(* IEC 61131-3 sources: STAR-PLC-Agent/results/raw/batch_fresh_20261114/PUB007/functional/attempt_0001, 1 file *)

(* ---- test_program.st ---- *)
PROGRAM PLC_PRG
VAR
 BenchStep : UDINT := 0;
 BenchCalls : UDINT := 0;
 BenchDone : BOOL := FALSE;
 BenchUut0 : FB_Task;
 BenchUut1 : FB_Task;
 BenchUut2 : FB_Task;
 BenchUut3 : FB_Task;
 BenchUut4 : FB_Task;
 BenchUut5 : FB_Task;
 BenchUut6 : FB_Task;
 Binding_0_pumpGroup : ARRAY[1..5] OF ST_Pump;
 Binding_1_pumpGroup : ARRAY[1..5] OF ST_Pump;
 Binding_2_pumpGroup : ARRAY[1..5] OF ST_Pump;
 Binding_3_pumpGroup : ARRAY[1..5] OF ST_Pump;
 Binding_4_pumpGroup : ARRAY[1..5] OF ST_Pump;
 Binding_5_pumpGroup : ARRAY[1..5] OF ST_Pump;
 Binding_6_pumpGroup : ARRAY[1..5] OF ST_Pump;
 TraceIn_mode : ARRAY[0..29] OF BOOL;
 TraceIn_start : ARRAY[0..29] OF BOOL;
 TraceIn_stop : ARRAY[0..29] OF BOOL;
 TraceOut_pumpGroup_1_priority : ARRAY[0..29] OF INT;
 TraceOut_pumpGroup_1_selection : ARRAY[0..29] OF BOOL;
 TraceOut_pumpGroup_1_RunComd : ARRAY[0..29] OF BOOL;
 TraceOut_pumpGroup_2_priority : ARRAY[0..29] OF INT;
 TraceOut_pumpGroup_2_selection : ARRAY[0..29] OF BOOL;
 TraceOut_pumpGroup_2_RunComd : ARRAY[0..29] OF BOOL;
 TraceOut_pumpGroup_3_priority : ARRAY[0..29] OF INT;
 TraceOut_pumpGroup_3_selection : ARRAY[0..29] OF BOOL;
 TraceOut_pumpGroup_3_RunComd : ARRAY[0..29] OF BOOL;
 TraceOut_pumpGroup_4_priority : ARRAY[0..29] OF INT;
 TraceOut_pumpGroup_4_selection : ARRAY[0..29] OF BOOL;
 TraceOut_pumpGroup_4_RunComd : ARRAY[0..29] OF BOOL;
 TraceOut_pumpGroup_5_priority : ARRAY[0..29] OF INT;
 TraceOut_pumpGroup_5_selection : ARRAY[0..29] OF BOOL;
 TraceOut_pumpGroup_5_RunComd : ARRAY[0..29] OF BOOL;
END_VAR

IF NOT BenchDone THEN
 CASE BenchStep OF
 0:
   Binding_0_pumpGroup[1].priority := INT#10;
   Binding_0_pumpGroup[1].selection := TRUE;
   Binding_0_pumpGroup[1].RunComd := FALSE;
   Binding_0_pumpGroup[2].priority := INT#20;
   Binding_0_pumpGroup[2].selection := FALSE;
   Binding_0_pumpGroup[2].RunComd := FALSE;
   Binding_0_pumpGroup[3].priority := INT#30;
   Binding_0_pumpGroup[3].selection := TRUE;
   Binding_0_pumpGroup[3].RunComd := FALSE;
   Binding_0_pumpGroup[4].priority := INT#40;
   Binding_0_pumpGroup[4].selection := FALSE;
   Binding_0_pumpGroup[4].RunComd := FALSE;
   Binding_0_pumpGroup[5].priority := INT#50;
   Binding_0_pumpGroup[5].selection := FALSE;
   Binding_0_pumpGroup[5].RunComd := FALSE;
   BenchUut0.mode := FALSE;
   BenchUut0.start := TRUE;
   BenchUut0.stop := FALSE;
   TraceIn_mode[0] := BenchUut0.mode;
   TraceIn_start[0] := BenchUut0.start;
   TraceIn_stop[0] := BenchUut0.stop;
   BenchUut0(pumpGroup := Binding_0_pumpGroup);
   TraceOut_pumpGroup_1_priority[0] := Binding_0_pumpGroup[1].priority;
   TraceOut_pumpGroup_1_selection[0] := Binding_0_pumpGroup[1].selection;
   TraceOut_pumpGroup_1_RunComd[0] := Binding_0_pumpGroup[1].RunComd;
   TraceOut_pumpGroup_2_priority[0] := Binding_0_pumpGroup[2].priority;
   TraceOut_pumpGroup_2_selection[0] := Binding_0_pumpGroup[2].selection;
   TraceOut_pumpGroup_2_RunComd[0] := Binding_0_pumpGroup[2].RunComd;
   TraceOut_pumpGroup_3_priority[0] := Binding_0_pumpGroup[3].priority;
   TraceOut_pumpGroup_3_selection[0] := Binding_0_pumpGroup[3].selection;
   TraceOut_pumpGroup_3_RunComd[0] := Binding_0_pumpGroup[3].RunComd;
   TraceOut_pumpGroup_4_priority[0] := Binding_0_pumpGroup[4].priority;
   TraceOut_pumpGroup_4_selection[0] := Binding_0_pumpGroup[4].selection;
   TraceOut_pumpGroup_4_RunComd[0] := Binding_0_pumpGroup[4].RunComd;
   TraceOut_pumpGroup_5_priority[0] := Binding_0_pumpGroup[5].priority;
   TraceOut_pumpGroup_5_selection[0] := Binding_0_pumpGroup[5].selection;
   TraceOut_pumpGroup_5_RunComd[0] := Binding_0_pumpGroup[5].RunComd;
   BenchCalls := BenchCalls + 1;
 1:
   Binding_0_pumpGroup[1].priority := INT#10;
   Binding_0_pumpGroup[1].selection := TRUE;
   Binding_0_pumpGroup[1].RunComd := TRUE;
   Binding_0_pumpGroup[2].priority := INT#20;
   Binding_0_pumpGroup[2].selection := FALSE;
   Binding_0_pumpGroup[2].RunComd := FALSE;
   Binding_0_pumpGroup[3].priority := INT#30;
   Binding_0_pumpGroup[3].selection := TRUE;
   Binding_0_pumpGroup[3].RunComd := TRUE;
   Binding_0_pumpGroup[4].priority := INT#40;
   Binding_0_pumpGroup[4].selection := FALSE;
   Binding_0_pumpGroup[4].RunComd := FALSE;
   Binding_0_pumpGroup[5].priority := INT#50;
   Binding_0_pumpGroup[5].selection := FALSE;
   Binding_0_pumpGroup[5].RunComd := FALSE;
   BenchUut0.mode := FALSE;
   BenchUut0.start := FALSE;
   BenchUut0.stop := FALSE;
   TraceIn_mode[1] := BenchUut0.mode;
   TraceIn_start[1] := BenchUut0.start;
   TraceIn_stop[1] := BenchUut0.stop;
   BenchUut0(pumpGroup := Binding_0_pumpGroup);
   TraceOut_pumpGroup_1_priority[1] := Binding_0_pumpGroup[1].priority;
   TraceOut_pumpGroup_1_selection[1] := Binding_0_pumpGroup[1].selection;
   TraceOut_pumpGroup_1_RunComd[1] := Binding_0_pumpGroup[1].RunComd;
   TraceOut_pumpGroup_2_priority[1] := Binding_0_pumpGroup[2].priority;
   TraceOut_pumpGroup_2_selection[1] := Binding_0_pumpGroup[2].selection;
   TraceOut_pumpGroup_2_RunComd[1] := Binding_0_pumpGroup[2].RunComd;
   TraceOut_pumpGroup_3_priority[1] := Binding_0_pumpGroup[3].priority;
   TraceOut_pumpGroup_3_selection[1] := Binding_0_pumpGroup[3].selection;
   TraceOut_pumpGroup_3_RunComd[1] := Binding_0_pumpGroup[3].RunComd;
   TraceOut_pumpGroup_4_priority[1] := Binding_0_pumpGroup[4].priority;
   TraceOut_pumpGroup_4_selection[1] := Binding_0_pumpGroup[4].selection;
   TraceOut_pumpGroup_4_RunComd[1] := Binding_0_pumpGroup[4].RunComd;
   TraceOut_pumpGroup_5_priority[1] := Binding_0_pumpGroup[5].priority;
   TraceOut_pumpGroup_5_selection[1] := Binding_0_pumpGroup[5].selection;
   TraceOut_pumpGroup_5_RunComd[1] := Binding_0_pumpGroup[5].RunComd;
   BenchCalls := BenchCalls + 1;
 2:
   Binding_0_pumpGroup[1].priority := INT#10;
   Binding_0_pumpGroup[1].selection := TRUE;
   Binding_0_pumpGroup[1].RunComd := TRUE;
   Binding_0_pumpGroup[2].priority := INT#20;
   Binding_0_pumpGroup[2].selection := FALSE;
   Binding_0_pumpGroup[2].RunComd := FALSE;
   Binding_0_pumpGroup[3].priority := INT#30;
   Binding_0_pumpGroup[3].selection := TRUE;
   Binding_0_pumpGroup[3].RunComd := TRUE;
   Binding_0_pumpGroup[4].priority := INT#40;
   Binding_0_pumpGroup[4].selection := FALSE;
   Binding_0_pumpGroup[4].RunComd := FALSE;
   Binding_0_pumpGroup[5].priority := INT#50;
   Binding_0_pumpGroup[5].selection := FALSE;
   Binding_0_pumpGroup[5].RunComd := FALSE;
   BenchUut0.mode := FALSE;
   BenchUut0.start := TRUE;
   BenchUut0.stop := TRUE;
   TraceIn_mode[2] := BenchUut0.mode;
   TraceIn_start[2] := BenchUut0.start;
   TraceIn_stop[2] := BenchUut0.stop;
   BenchUut0(pumpGroup := Binding_0_pumpGroup);
   TraceOut_pumpGroup_1_priority[2] := Binding_0_pumpGroup[1].priority;
   TraceOut_pumpGroup_1_selection[2] := Binding_0_pumpGroup[1].selection;
   TraceOut_pumpGroup_1_RunComd[2] := Binding_0_pumpGroup[1].RunComd;
   TraceOut_pumpGroup_2_priority[2] := Binding_0_pumpGroup[2].priority;
   TraceOut_pumpGroup_2_selection[2] := Binding_0_pumpGroup[2].selection;
   TraceOut_pumpGroup_2_RunComd[2] := Binding_0_pumpGroup[2].RunComd;
   TraceOut_pumpGroup_3_priority[2] := Binding_0_pumpGroup[3].priority;
   TraceOut_pumpGroup_3_selection[2] := Binding_0_pumpGroup[3].selection;
   TraceOut_pumpGroup_3_RunComd[2] := Binding_0_pumpGroup[3].RunComd;
   TraceOut_pumpGroup_4_priority[2] := Binding_0_pumpGroup[4].priority;
   TraceOut_pumpGroup_4_selection[2] := Binding_0_pumpGroup[4].selection;
   TraceOut_pumpGroup_4_RunComd[2] := Binding_0_pumpGroup[4].RunComd;
   TraceOut_pumpGroup_5_priority[2] := Binding_0_pumpGroup[5].priority;
   TraceOut_pumpGroup_5_selection[2] := Binding_0_pumpGroup[5].selection;
   TraceOut_pumpGroup_5_RunComd[2] := Binding_0_pumpGroup[5].RunComd;
   BenchCalls := BenchCalls + 1;
 3:
   Binding_1_pumpGroup[1].priority := INT#10;
   Binding_1_pumpGroup[1].selection := TRUE;
   Binding_1_pumpGroup[1].RunComd := FALSE;
   Binding_1_pumpGroup[2].priority := INT#20;
   Binding_1_pumpGroup[2].selection := FALSE;
   Binding_1_pumpGroup[2].RunComd := FALSE;
   Binding_1_pumpGroup[3].priority := INT#30;
   Binding_1_pumpGroup[3].selection := TRUE;
   Binding_1_pumpGroup[3].RunComd := FALSE;
   Binding_1_pumpGroup[4].priority := INT#40;
   Binding_1_pumpGroup[4].selection := FALSE;
   Binding_1_pumpGroup[4].RunComd := FALSE;
   Binding_1_pumpGroup[5].priority := INT#50;
   Binding_1_pumpGroup[5].selection := FALSE;
   Binding_1_pumpGroup[5].RunComd := FALSE;
   BenchUut1.mode := TRUE;
   BenchUut1.start := TRUE;
   BenchUut1.stop := FALSE;
   TraceIn_mode[3] := BenchUut1.mode;
   TraceIn_start[3] := BenchUut1.start;
   TraceIn_stop[3] := BenchUut1.stop;
   BenchUut1(pumpGroup := Binding_1_pumpGroup);
   TraceOut_pumpGroup_1_priority[3] := Binding_1_pumpGroup[1].priority;
   TraceOut_pumpGroup_1_selection[3] := Binding_1_pumpGroup[1].selection;
   TraceOut_pumpGroup_1_RunComd[3] := Binding_1_pumpGroup[1].RunComd;
   TraceOut_pumpGroup_2_priority[3] := Binding_1_pumpGroup[2].priority;
   TraceOut_pumpGroup_2_selection[3] := Binding_1_pumpGroup[2].selection;
   TraceOut_pumpGroup_2_RunComd[3] := Binding_1_pumpGroup[2].RunComd;
   TraceOut_pumpGroup_3_priority[3] := Binding_1_pumpGroup[3].priority;
   TraceOut_pumpGroup_3_selection[3] := Binding_1_pumpGroup[3].selection;
   TraceOut_pumpGroup_3_RunComd[3] := Binding_1_pumpGroup[3].RunComd;
   TraceOut_pumpGroup_4_priority[3] := Binding_1_pumpGroup[4].priority;
   TraceOut_pumpGroup_4_selection[3] := Binding_1_pumpGroup[4].selection;
   TraceOut_pumpGroup_4_RunComd[3] := Binding_1_pumpGroup[4].RunComd;
   TraceOut_pumpGroup_5_priority[3] := Binding_1_pumpGroup[5].priority;
   TraceOut_pumpGroup_5_selection[3] := Binding_1_pumpGroup[5].selection;
   TraceOut_pumpGroup_5_RunComd[3] := Binding_1_pumpGroup[5].RunComd;
   BenchCalls := BenchCalls + 1;
 4:
   Binding_1_pumpGroup[1].priority := INT#5;
   Binding_1_pumpGroup[1].selection := TRUE;
   Binding_1_pumpGroup[1].RunComd := FALSE;
   Binding_1_pumpGroup[2].priority := INT#5;
   Binding_1_pumpGroup[2].selection := FALSE;
   Binding_1_pumpGroup[2].RunComd := FALSE;
   Binding_1_pumpGroup[3].priority := INT#5;
   Binding_1_pumpGroup[3].selection := TRUE;
   Binding_1_pumpGroup[3].RunComd := TRUE;
   Binding_1_pumpGroup[4].priority := INT#5;
   Binding_1_pumpGroup[4].selection := FALSE;
   Binding_1_pumpGroup[4].RunComd := TRUE;
   Binding_1_pumpGroup[5].priority := INT#5;
   Binding_1_pumpGroup[5].selection := FALSE;
   Binding_1_pumpGroup[5].RunComd := TRUE;
   BenchUut1.mode := TRUE;
   BenchUut1.start := TRUE;
   BenchUut1.stop := FALSE;
   TraceIn_mode[4] := BenchUut1.mode;
   TraceIn_start[4] := BenchUut1.start;
   TraceIn_stop[4] := BenchUut1.stop;
   BenchUut1(pumpGroup := Binding_1_pumpGroup);
   TraceOut_pumpGroup_1_priority[4] := Binding_1_pumpGroup[1].priority;
   TraceOut_pumpGroup_1_selection[4] := Binding_1_pumpGroup[1].selection;
   TraceOut_pumpGroup_1_RunComd[4] := Binding_1_pumpGroup[1].RunComd;
   TraceOut_pumpGroup_2_priority[4] := Binding_1_pumpGroup[2].priority;
   TraceOut_pumpGroup_2_selection[4] := Binding_1_pumpGroup[2].selection;
   TraceOut_pumpGroup_2_RunComd[4] := Binding_1_pumpGroup[2].RunComd;
   TraceOut_pumpGroup_3_priority[4] := Binding_1_pumpGroup[3].priority;
   TraceOut_pumpGroup_3_selection[4] := Binding_1_pumpGroup[3].selection;
   TraceOut_pumpGroup_3_RunComd[4] := Binding_1_pumpGroup[3].RunComd;
   TraceOut_pumpGroup_4_priority[4] := Binding_1_pumpGroup[4].priority;
   TraceOut_pumpGroup_4_selection[4] := Binding_1_pumpGroup[4].selection;
   TraceOut_pumpGroup_4_RunComd[4] := Binding_1_pumpGroup[4].RunComd;
   TraceOut_pumpGroup_5_priority[4] := Binding_1_pumpGroup[5].priority;
   TraceOut_pumpGroup_5_selection[4] := Binding_1_pumpGroup[5].selection;
   TraceOut_pumpGroup_5_RunComd[4] := Binding_1_pumpGroup[5].RunComd;
   BenchCalls := BenchCalls + 1;
 5:
   Binding_1_pumpGroup[1].priority := INT#-3;
   Binding_1_pumpGroup[1].selection := TRUE;
   Binding_1_pumpGroup[1].RunComd := TRUE;
   Binding_1_pumpGroup[2].priority := INT#0;
   Binding_1_pumpGroup[2].selection := FALSE;
   Binding_1_pumpGroup[2].RunComd := TRUE;
   Binding_1_pumpGroup[3].priority := INT#-1;
   Binding_1_pumpGroup[3].selection := TRUE;
   Binding_1_pumpGroup[3].RunComd := TRUE;
   Binding_1_pumpGroup[4].priority := INT#-2;
   Binding_1_pumpGroup[4].selection := FALSE;
   Binding_1_pumpGroup[4].RunComd := FALSE;
   Binding_1_pumpGroup[5].priority := INT#4;
   Binding_1_pumpGroup[5].selection := FALSE;
   Binding_1_pumpGroup[5].RunComd := FALSE;
   BenchUut1.mode := TRUE;
   BenchUut1.start := TRUE;
   BenchUut1.stop := FALSE;
   TraceIn_mode[5] := BenchUut1.mode;
   TraceIn_start[5] := BenchUut1.start;
   TraceIn_stop[5] := BenchUut1.stop;
   BenchUut1(pumpGroup := Binding_1_pumpGroup);
   TraceOut_pumpGroup_1_priority[5] := Binding_1_pumpGroup[1].priority;
   TraceOut_pumpGroup_1_selection[5] := Binding_1_pumpGroup[1].selection;
   TraceOut_pumpGroup_1_RunComd[5] := Binding_1_pumpGroup[1].RunComd;
   TraceOut_pumpGroup_2_priority[5] := Binding_1_pumpGroup[2].priority;
   TraceOut_pumpGroup_2_selection[5] := Binding_1_pumpGroup[2].selection;
   TraceOut_pumpGroup_2_RunComd[5] := Binding_1_pumpGroup[2].RunComd;
   TraceOut_pumpGroup_3_priority[5] := Binding_1_pumpGroup[3].priority;
   TraceOut_pumpGroup_3_selection[5] := Binding_1_pumpGroup[3].selection;
   TraceOut_pumpGroup_3_RunComd[5] := Binding_1_pumpGroup[3].RunComd;
   TraceOut_pumpGroup_4_priority[5] := Binding_1_pumpGroup[4].priority;
   TraceOut_pumpGroup_4_selection[5] := Binding_1_pumpGroup[4].selection;
   TraceOut_pumpGroup_4_RunComd[5] := Binding_1_pumpGroup[4].RunComd;
   TraceOut_pumpGroup_5_priority[5] := Binding_1_pumpGroup[5].priority;
   TraceOut_pumpGroup_5_selection[5] := Binding_1_pumpGroup[5].selection;
   TraceOut_pumpGroup_5_RunComd[5] := Binding_1_pumpGroup[5].RunComd;
   BenchCalls := BenchCalls + 1;
 6:
   Binding_2_pumpGroup[1].priority := INT#1;
   Binding_2_pumpGroup[1].selection := FALSE;
   Binding_2_pumpGroup[1].RunComd := FALSE;
   Binding_2_pumpGroup[2].priority := INT#1;
   Binding_2_pumpGroup[2].selection := FALSE;
   Binding_2_pumpGroup[2].RunComd := FALSE;
   Binding_2_pumpGroup[3].priority := INT#1;
   Binding_2_pumpGroup[3].selection := FALSE;
   Binding_2_pumpGroup[3].RunComd := FALSE;
   Binding_2_pumpGroup[4].priority := INT#1;
   Binding_2_pumpGroup[4].selection := FALSE;
   Binding_2_pumpGroup[4].RunComd := FALSE;
   Binding_2_pumpGroup[5].priority := INT#1;
   Binding_2_pumpGroup[5].selection := FALSE;
   Binding_2_pumpGroup[5].RunComd := FALSE;
   BenchUut2.mode := TRUE;
   BenchUut2.start := TRUE;
   BenchUut2.stop := FALSE;
   TraceIn_mode[6] := BenchUut2.mode;
   TraceIn_start[6] := BenchUut2.start;
   TraceIn_stop[6] := BenchUut2.stop;
   BenchUut2(pumpGroup := Binding_2_pumpGroup);
   TraceOut_pumpGroup_1_priority[6] := Binding_2_pumpGroup[1].priority;
   TraceOut_pumpGroup_1_selection[6] := Binding_2_pumpGroup[1].selection;
   TraceOut_pumpGroup_1_RunComd[6] := Binding_2_pumpGroup[1].RunComd;
   TraceOut_pumpGroup_2_priority[6] := Binding_2_pumpGroup[2].priority;
   TraceOut_pumpGroup_2_selection[6] := Binding_2_pumpGroup[2].selection;
   TraceOut_pumpGroup_2_RunComd[6] := Binding_2_pumpGroup[2].RunComd;
   TraceOut_pumpGroup_3_priority[6] := Binding_2_pumpGroup[3].priority;
   TraceOut_pumpGroup_3_selection[6] := Binding_2_pumpGroup[3].selection;
   TraceOut_pumpGroup_3_RunComd[6] := Binding_2_pumpGroup[3].RunComd;
   TraceOut_pumpGroup_4_priority[6] := Binding_2_pumpGroup[4].priority;
   TraceOut_pumpGroup_4_selection[6] := Binding_2_pumpGroup[4].selection;
   TraceOut_pumpGroup_4_RunComd[6] := Binding_2_pumpGroup[4].RunComd;
   TraceOut_pumpGroup_5_priority[6] := Binding_2_pumpGroup[5].priority;
   TraceOut_pumpGroup_5_selection[6] := Binding_2_pumpGroup[5].selection;
   TraceOut_pumpGroup_5_RunComd[6] := Binding_2_pumpGroup[5].RunComd;
   BenchCalls := BenchCalls + 1;
 7:
   Binding_2_pumpGroup[1].priority := INT#1;
   Binding_2_pumpGroup[1].selection := FALSE;
   Binding_2_pumpGroup[1].RunComd := TRUE;
   Binding_2_pumpGroup[2].priority := INT#2;
   Binding_2_pumpGroup[2].selection := FALSE;
   Binding_2_pumpGroup[2].RunComd := TRUE;
   Binding_2_pumpGroup[3].priority := INT#3;
   Binding_2_pumpGroup[3].selection := FALSE;
   Binding_2_pumpGroup[3].RunComd := TRUE;
   Binding_2_pumpGroup[4].priority := INT#4;
   Binding_2_pumpGroup[4].selection := FALSE;
   Binding_2_pumpGroup[4].RunComd := FALSE;
   Binding_2_pumpGroup[5].priority := INT#5;
   Binding_2_pumpGroup[5].selection := FALSE;
   Binding_2_pumpGroup[5].RunComd := FALSE;
   BenchUut2.mode := TRUE;
   BenchUut2.start := FALSE;
   BenchUut2.stop := FALSE;
   TraceIn_mode[7] := BenchUut2.mode;
   TraceIn_start[7] := BenchUut2.start;
   TraceIn_stop[7] := BenchUut2.stop;
   BenchUut2(pumpGroup := Binding_2_pumpGroup);
   TraceOut_pumpGroup_1_priority[7] := Binding_2_pumpGroup[1].priority;
   TraceOut_pumpGroup_1_selection[7] := Binding_2_pumpGroup[1].selection;
   TraceOut_pumpGroup_1_RunComd[7] := Binding_2_pumpGroup[1].RunComd;
   TraceOut_pumpGroup_2_priority[7] := Binding_2_pumpGroup[2].priority;
   TraceOut_pumpGroup_2_selection[7] := Binding_2_pumpGroup[2].selection;
   TraceOut_pumpGroup_2_RunComd[7] := Binding_2_pumpGroup[2].RunComd;
   TraceOut_pumpGroup_3_priority[7] := Binding_2_pumpGroup[3].priority;
   TraceOut_pumpGroup_3_selection[7] := Binding_2_pumpGroup[3].selection;
   TraceOut_pumpGroup_3_RunComd[7] := Binding_2_pumpGroup[3].RunComd;
   TraceOut_pumpGroup_4_priority[7] := Binding_2_pumpGroup[4].priority;
   TraceOut_pumpGroup_4_selection[7] := Binding_2_pumpGroup[4].selection;
   TraceOut_pumpGroup_4_RunComd[7] := Binding_2_pumpGroup[4].RunComd;
   TraceOut_pumpGroup_5_priority[7] := Binding_2_pumpGroup[5].priority;
   TraceOut_pumpGroup_5_selection[7] := Binding_2_pumpGroup[5].selection;
   TraceOut_pumpGroup_5_RunComd[7] := Binding_2_pumpGroup[5].RunComd;
   BenchCalls := BenchCalls + 1;
 8:
   Binding_2_pumpGroup[1].priority := INT#1;
   Binding_2_pumpGroup[1].selection := FALSE;
   Binding_2_pumpGroup[1].RunComd := TRUE;
   Binding_2_pumpGroup[2].priority := INT#2;
   Binding_2_pumpGroup[2].selection := FALSE;
   Binding_2_pumpGroup[2].RunComd := TRUE;
   Binding_2_pumpGroup[3].priority := INT#3;
   Binding_2_pumpGroup[3].selection := FALSE;
   Binding_2_pumpGroup[3].RunComd := TRUE;
   Binding_2_pumpGroup[4].priority := INT#4;
   Binding_2_pumpGroup[4].selection := FALSE;
   Binding_2_pumpGroup[4].RunComd := FALSE;
   Binding_2_pumpGroup[5].priority := INT#5;
   Binding_2_pumpGroup[5].selection := FALSE;
   Binding_2_pumpGroup[5].RunComd := FALSE;
   BenchUut2.mode := TRUE;
   BenchUut2.start := TRUE;
   BenchUut2.stop := FALSE;
   TraceIn_mode[8] := BenchUut2.mode;
   TraceIn_start[8] := BenchUut2.start;
   TraceIn_stop[8] := BenchUut2.stop;
   BenchUut2(pumpGroup := Binding_2_pumpGroup);
   TraceOut_pumpGroup_1_priority[8] := Binding_2_pumpGroup[1].priority;
   TraceOut_pumpGroup_1_selection[8] := Binding_2_pumpGroup[1].selection;
   TraceOut_pumpGroup_1_RunComd[8] := Binding_2_pumpGroup[1].RunComd;
   TraceOut_pumpGroup_2_priority[8] := Binding_2_pumpGroup[2].priority;
   TraceOut_pumpGroup_2_selection[8] := Binding_2_pumpGroup[2].selection;
   TraceOut_pumpGroup_2_RunComd[8] := Binding_2_pumpGroup[2].RunComd;
   TraceOut_pumpGroup_3_priority[8] := Binding_2_pumpGroup[3].priority;
   TraceOut_pumpGroup_3_selection[8] := Binding_2_pumpGroup[3].selection;
   TraceOut_pumpGroup_3_RunComd[8] := Binding_2_pumpGroup[3].RunComd;
   TraceOut_pumpGroup_4_priority[8] := Binding_2_pumpGroup[4].priority;
   TraceOut_pumpGroup_4_selection[8] := Binding_2_pumpGroup[4].selection;
   TraceOut_pumpGroup_4_RunComd[8] := Binding_2_pumpGroup[4].RunComd;
   TraceOut_pumpGroup_5_priority[8] := Binding_2_pumpGroup[5].priority;
   TraceOut_pumpGroup_5_selection[8] := Binding_2_pumpGroup[5].selection;
   TraceOut_pumpGroup_5_RunComd[8] := Binding_2_pumpGroup[5].RunComd;
   BenchCalls := BenchCalls + 1;
 9:
   Binding_2_pumpGroup[1].priority := INT#1;
   Binding_2_pumpGroup[1].selection := FALSE;
   Binding_2_pumpGroup[1].RunComd := FALSE;
   Binding_2_pumpGroup[2].priority := INT#1;
   Binding_2_pumpGroup[2].selection := FALSE;
   Binding_2_pumpGroup[2].RunComd := FALSE;
   Binding_2_pumpGroup[3].priority := INT#1;
   Binding_2_pumpGroup[3].selection := FALSE;
   Binding_2_pumpGroup[3].RunComd := TRUE;
   Binding_2_pumpGroup[4].priority := INT#1;
   Binding_2_pumpGroup[4].selection := FALSE;
   Binding_2_pumpGroup[4].RunComd := TRUE;
   Binding_2_pumpGroup[5].priority := INT#1;
   Binding_2_pumpGroup[5].selection := FALSE;
   Binding_2_pumpGroup[5].RunComd := TRUE;
   BenchUut2.mode := TRUE;
   BenchUut2.start := TRUE;
   BenchUut2.stop := TRUE;
   TraceIn_mode[9] := BenchUut2.mode;
   TraceIn_start[9] := BenchUut2.start;
   TraceIn_stop[9] := BenchUut2.stop;
   BenchUut2(pumpGroup := Binding_2_pumpGroup);
   TraceOut_pumpGroup_1_priority[9] := Binding_2_pumpGroup[1].priority;
   TraceOut_pumpGroup_1_selection[9] := Binding_2_pumpGroup[1].selection;
   TraceOut_pumpGroup_1_RunComd[9] := Binding_2_pumpGroup[1].RunComd;
   TraceOut_pumpGroup_2_priority[9] := Binding_2_pumpGroup[2].priority;
   TraceOut_pumpGroup_2_selection[9] := Binding_2_pumpGroup[2].selection;
   TraceOut_pumpGroup_2_RunComd[9] := Binding_2_pumpGroup[2].RunComd;
   TraceOut_pumpGroup_3_priority[9] := Binding_2_pumpGroup[3].priority;
   TraceOut_pumpGroup_3_selection[9] := Binding_2_pumpGroup[3].selection;
   TraceOut_pumpGroup_3_RunComd[9] := Binding_2_pumpGroup[3].RunComd;
   TraceOut_pumpGroup_4_priority[9] := Binding_2_pumpGroup[4].priority;
   TraceOut_pumpGroup_4_selection[9] := Binding_2_pumpGroup[4].selection;
   TraceOut_pumpGroup_4_RunComd[9] := Binding_2_pumpGroup[4].RunComd;
   TraceOut_pumpGroup_5_priority[9] := Binding_2_pumpGroup[5].priority;
   TraceOut_pumpGroup_5_selection[9] := Binding_2_pumpGroup[5].selection;
   TraceOut_pumpGroup_5_RunComd[9] := Binding_2_pumpGroup[5].RunComd;
   BenchCalls := BenchCalls + 1;
 10:
   Binding_3_pumpGroup[1].priority := INT#1;
   Binding_3_pumpGroup[1].selection := TRUE;
   Binding_3_pumpGroup[1].RunComd := FALSE;
   Binding_3_pumpGroup[2].priority := INT#2;
   Binding_3_pumpGroup[2].selection := FALSE;
   Binding_3_pumpGroup[2].RunComd := FALSE;
   Binding_3_pumpGroup[3].priority := INT#3;
   Binding_3_pumpGroup[3].selection := TRUE;
   Binding_3_pumpGroup[3].RunComd := FALSE;
   Binding_3_pumpGroup[4].priority := INT#4;
   Binding_3_pumpGroup[4].selection := FALSE;
   Binding_3_pumpGroup[4].RunComd := FALSE;
   Binding_3_pumpGroup[5].priority := INT#5;
   Binding_3_pumpGroup[5].selection := TRUE;
   Binding_3_pumpGroup[5].RunComd := FALSE;
   BenchUut3.mode := FALSE;
   BenchUut3.start := TRUE;
   BenchUut3.stop := FALSE;
   TraceIn_mode[10] := BenchUut3.mode;
   TraceIn_start[10] := BenchUut3.start;
   TraceIn_stop[10] := BenchUut3.stop;
   BenchUut3(pumpGroup := Binding_3_pumpGroup);
   TraceOut_pumpGroup_1_priority[10] := Binding_3_pumpGroup[1].priority;
   TraceOut_pumpGroup_1_selection[10] := Binding_3_pumpGroup[1].selection;
   TraceOut_pumpGroup_1_RunComd[10] := Binding_3_pumpGroup[1].RunComd;
   TraceOut_pumpGroup_2_priority[10] := Binding_3_pumpGroup[2].priority;
   TraceOut_pumpGroup_2_selection[10] := Binding_3_pumpGroup[2].selection;
   TraceOut_pumpGroup_2_RunComd[10] := Binding_3_pumpGroup[2].RunComd;
   TraceOut_pumpGroup_3_priority[10] := Binding_3_pumpGroup[3].priority;
   TraceOut_pumpGroup_3_selection[10] := Binding_3_pumpGroup[3].selection;
   TraceOut_pumpGroup_3_RunComd[10] := Binding_3_pumpGroup[3].RunComd;
   TraceOut_pumpGroup_4_priority[10] := Binding_3_pumpGroup[4].priority;
   TraceOut_pumpGroup_4_selection[10] := Binding_3_pumpGroup[4].selection;
   TraceOut_pumpGroup_4_RunComd[10] := Binding_3_pumpGroup[4].RunComd;
   TraceOut_pumpGroup_5_priority[10] := Binding_3_pumpGroup[5].priority;
   TraceOut_pumpGroup_5_selection[10] := Binding_3_pumpGroup[5].selection;
   TraceOut_pumpGroup_5_RunComd[10] := Binding_3_pumpGroup[5].RunComd;
   BenchCalls := BenchCalls + 1;
 11:
   Binding_3_pumpGroup[1].priority := INT#100;
   Binding_3_pumpGroup[1].selection := FALSE;
   Binding_3_pumpGroup[1].RunComd := TRUE;
   Binding_3_pumpGroup[2].priority := INT#100;
   Binding_3_pumpGroup[2].selection := FALSE;
   Binding_3_pumpGroup[2].RunComd := FALSE;
   Binding_3_pumpGroup[3].priority := INT#5;
   Binding_3_pumpGroup[3].selection := FALSE;
   Binding_3_pumpGroup[3].RunComd := TRUE;
   Binding_3_pumpGroup[4].priority := INT#5;
   Binding_3_pumpGroup[4].selection := FALSE;
   Binding_3_pumpGroup[4].RunComd := FALSE;
   Binding_3_pumpGroup[5].priority := INT#5;
   Binding_3_pumpGroup[5].selection := FALSE;
   Binding_3_pumpGroup[5].RunComd := TRUE;
   BenchUut3.mode := TRUE;
   BenchUut3.start := FALSE;
   BenchUut3.stop := FALSE;
   TraceIn_mode[11] := BenchUut3.mode;
   TraceIn_start[11] := BenchUut3.start;
   TraceIn_stop[11] := BenchUut3.stop;
   BenchUut3(pumpGroup := Binding_3_pumpGroup);
   TraceOut_pumpGroup_1_priority[11] := Binding_3_pumpGroup[1].priority;
   TraceOut_pumpGroup_1_selection[11] := Binding_3_pumpGroup[1].selection;
   TraceOut_pumpGroup_1_RunComd[11] := Binding_3_pumpGroup[1].RunComd;
   TraceOut_pumpGroup_2_priority[11] := Binding_3_pumpGroup[2].priority;
   TraceOut_pumpGroup_2_selection[11] := Binding_3_pumpGroup[2].selection;
   TraceOut_pumpGroup_2_RunComd[11] := Binding_3_pumpGroup[2].RunComd;
   TraceOut_pumpGroup_3_priority[11] := Binding_3_pumpGroup[3].priority;
   TraceOut_pumpGroup_3_selection[11] := Binding_3_pumpGroup[3].selection;
   TraceOut_pumpGroup_3_RunComd[11] := Binding_3_pumpGroup[3].RunComd;
   TraceOut_pumpGroup_4_priority[11] := Binding_3_pumpGroup[4].priority;
   TraceOut_pumpGroup_4_selection[11] := Binding_3_pumpGroup[4].selection;
   TraceOut_pumpGroup_4_RunComd[11] := Binding_3_pumpGroup[4].RunComd;
   TraceOut_pumpGroup_5_priority[11] := Binding_3_pumpGroup[5].priority;
   TraceOut_pumpGroup_5_selection[11] := Binding_3_pumpGroup[5].selection;
   TraceOut_pumpGroup_5_RunComd[11] := Binding_3_pumpGroup[5].RunComd;
   BenchCalls := BenchCalls + 1;
 12:
   Binding_3_pumpGroup[1].priority := INT#100;
   Binding_3_pumpGroup[1].selection := FALSE;
   Binding_3_pumpGroup[1].RunComd := TRUE;
   Binding_3_pumpGroup[2].priority := INT#100;
   Binding_3_pumpGroup[2].selection := FALSE;
   Binding_3_pumpGroup[2].RunComd := FALSE;
   Binding_3_pumpGroup[3].priority := INT#5;
   Binding_3_pumpGroup[3].selection := FALSE;
   Binding_3_pumpGroup[3].RunComd := TRUE;
   Binding_3_pumpGroup[4].priority := INT#5;
   Binding_3_pumpGroup[4].selection := FALSE;
   Binding_3_pumpGroup[4].RunComd := FALSE;
   Binding_3_pumpGroup[5].priority := INT#5;
   Binding_3_pumpGroup[5].selection := FALSE;
   Binding_3_pumpGroup[5].RunComd := TRUE;
   BenchUut3.mode := TRUE;
   BenchUut3.start := TRUE;
   BenchUut3.stop := FALSE;
   TraceIn_mode[12] := BenchUut3.mode;
   TraceIn_start[12] := BenchUut3.start;
   TraceIn_stop[12] := BenchUut3.stop;
   BenchUut3(pumpGroup := Binding_3_pumpGroup);
   TraceOut_pumpGroup_1_priority[12] := Binding_3_pumpGroup[1].priority;
   TraceOut_pumpGroup_1_selection[12] := Binding_3_pumpGroup[1].selection;
   TraceOut_pumpGroup_1_RunComd[12] := Binding_3_pumpGroup[1].RunComd;
   TraceOut_pumpGroup_2_priority[12] := Binding_3_pumpGroup[2].priority;
   TraceOut_pumpGroup_2_selection[12] := Binding_3_pumpGroup[2].selection;
   TraceOut_pumpGroup_2_RunComd[12] := Binding_3_pumpGroup[2].RunComd;
   TraceOut_pumpGroup_3_priority[12] := Binding_3_pumpGroup[3].priority;
   TraceOut_pumpGroup_3_selection[12] := Binding_3_pumpGroup[3].selection;
   TraceOut_pumpGroup_3_RunComd[12] := Binding_3_pumpGroup[3].RunComd;
   TraceOut_pumpGroup_4_priority[12] := Binding_3_pumpGroup[4].priority;
   TraceOut_pumpGroup_4_selection[12] := Binding_3_pumpGroup[4].selection;
   TraceOut_pumpGroup_4_RunComd[12] := Binding_3_pumpGroup[4].RunComd;
   TraceOut_pumpGroup_5_priority[12] := Binding_3_pumpGroup[5].priority;
   TraceOut_pumpGroup_5_selection[12] := Binding_3_pumpGroup[5].selection;
   TraceOut_pumpGroup_5_RunComd[12] := Binding_3_pumpGroup[5].RunComd;
   BenchCalls := BenchCalls + 1;
 13:
   Binding_3_pumpGroup[1].priority := INT#100;
   Binding_3_pumpGroup[1].selection := FALSE;
   Binding_3_pumpGroup[1].RunComd := TRUE;
   Binding_3_pumpGroup[2].priority := INT#100;
   Binding_3_pumpGroup[2].selection := FALSE;
   Binding_3_pumpGroup[2].RunComd := TRUE;
   Binding_3_pumpGroup[3].priority := INT#5;
   Binding_3_pumpGroup[3].selection := FALSE;
   Binding_3_pumpGroup[3].RunComd := TRUE;
   Binding_3_pumpGroup[4].priority := INT#5;
   Binding_3_pumpGroup[4].selection := FALSE;
   Binding_3_pumpGroup[4].RunComd := FALSE;
   Binding_3_pumpGroup[5].priority := INT#5;
   Binding_3_pumpGroup[5].selection := FALSE;
   Binding_3_pumpGroup[5].RunComd := FALSE;
   BenchUut3.mode := TRUE;
   BenchUut3.start := TRUE;
   BenchUut3.stop := TRUE;
   TraceIn_mode[13] := BenchUut3.mode;
   TraceIn_start[13] := BenchUut3.start;
   TraceIn_stop[13] := BenchUut3.stop;
   BenchUut3(pumpGroup := Binding_3_pumpGroup);
   TraceOut_pumpGroup_1_priority[13] := Binding_3_pumpGroup[1].priority;
   TraceOut_pumpGroup_1_selection[13] := Binding_3_pumpGroup[1].selection;
   TraceOut_pumpGroup_1_RunComd[13] := Binding_3_pumpGroup[1].RunComd;
   TraceOut_pumpGroup_2_priority[13] := Binding_3_pumpGroup[2].priority;
   TraceOut_pumpGroup_2_selection[13] := Binding_3_pumpGroup[2].selection;
   TraceOut_pumpGroup_2_RunComd[13] := Binding_3_pumpGroup[2].RunComd;
   TraceOut_pumpGroup_3_priority[13] := Binding_3_pumpGroup[3].priority;
   TraceOut_pumpGroup_3_selection[13] := Binding_3_pumpGroup[3].selection;
   TraceOut_pumpGroup_3_RunComd[13] := Binding_3_pumpGroup[3].RunComd;
   TraceOut_pumpGroup_4_priority[13] := Binding_3_pumpGroup[4].priority;
   TraceOut_pumpGroup_4_selection[13] := Binding_3_pumpGroup[4].selection;
   TraceOut_pumpGroup_4_RunComd[13] := Binding_3_pumpGroup[4].RunComd;
   TraceOut_pumpGroup_5_priority[13] := Binding_3_pumpGroup[5].priority;
   TraceOut_pumpGroup_5_selection[13] := Binding_3_pumpGroup[5].selection;
   TraceOut_pumpGroup_5_RunComd[13] := Binding_3_pumpGroup[5].RunComd;
   BenchCalls := BenchCalls + 1;
 14:
   Binding_3_pumpGroup[1].priority := INT#-32768;
   Binding_3_pumpGroup[1].selection := FALSE;
   Binding_3_pumpGroup[1].RunComd := FALSE;
   Binding_3_pumpGroup[2].priority := INT#32767;
   Binding_3_pumpGroup[2].selection := FALSE;
   Binding_3_pumpGroup[2].RunComd := FALSE;
   Binding_3_pumpGroup[3].priority := INT#0;
   Binding_3_pumpGroup[3].selection := FALSE;
   Binding_3_pumpGroup[3].RunComd := FALSE;
   Binding_3_pumpGroup[4].priority := INT#32766;
   Binding_3_pumpGroup[4].selection := FALSE;
   Binding_3_pumpGroup[4].RunComd := FALSE;
   Binding_3_pumpGroup[5].priority := INT#-1;
   Binding_3_pumpGroup[5].selection := FALSE;
   Binding_3_pumpGroup[5].RunComd := FALSE;
   BenchUut3.mode := TRUE;
   BenchUut3.start := TRUE;
   BenchUut3.stop := FALSE;
   TraceIn_mode[14] := BenchUut3.mode;
   TraceIn_start[14] := BenchUut3.start;
   TraceIn_stop[14] := BenchUut3.stop;
   BenchUut3(pumpGroup := Binding_3_pumpGroup);
   TraceOut_pumpGroup_1_priority[14] := Binding_3_pumpGroup[1].priority;
   TraceOut_pumpGroup_1_selection[14] := Binding_3_pumpGroup[1].selection;
   TraceOut_pumpGroup_1_RunComd[14] := Binding_3_pumpGroup[1].RunComd;
   TraceOut_pumpGroup_2_priority[14] := Binding_3_pumpGroup[2].priority;
   TraceOut_pumpGroup_2_selection[14] := Binding_3_pumpGroup[2].selection;
   TraceOut_pumpGroup_2_RunComd[14] := Binding_3_pumpGroup[2].RunComd;
   TraceOut_pumpGroup_3_priority[14] := Binding_3_pumpGroup[3].priority;
   TraceOut_pumpGroup_3_selection[14] := Binding_3_pumpGroup[3].selection;
   TraceOut_pumpGroup_3_RunComd[14] := Binding_3_pumpGroup[3].RunComd;
   TraceOut_pumpGroup_4_priority[14] := Binding_3_pumpGroup[4].priority;
   TraceOut_pumpGroup_4_selection[14] := Binding_3_pumpGroup[4].selection;
   TraceOut_pumpGroup_4_RunComd[14] := Binding_3_pumpGroup[4].RunComd;
   TraceOut_pumpGroup_5_priority[14] := Binding_3_pumpGroup[5].priority;
   TraceOut_pumpGroup_5_selection[14] := Binding_3_pumpGroup[5].selection;
   TraceOut_pumpGroup_5_RunComd[14] := Binding_3_pumpGroup[5].RunComd;
   BenchCalls := BenchCalls + 1;
 15:
   Binding_4_pumpGroup[1].priority := INT#10;
   Binding_4_pumpGroup[1].selection := TRUE;
   Binding_4_pumpGroup[1].RunComd := FALSE;
   Binding_4_pumpGroup[2].priority := INT#20;
   Binding_4_pumpGroup[2].selection := FALSE;
   Binding_4_pumpGroup[2].RunComd := FALSE;
   Binding_4_pumpGroup[3].priority := INT#30;
   Binding_4_pumpGroup[3].selection := TRUE;
   Binding_4_pumpGroup[3].RunComd := FALSE;
   Binding_4_pumpGroup[4].priority := INT#40;
   Binding_4_pumpGroup[4].selection := FALSE;
   Binding_4_pumpGroup[4].RunComd := FALSE;
   Binding_4_pumpGroup[5].priority := INT#50;
   Binding_4_pumpGroup[5].selection := FALSE;
   Binding_4_pumpGroup[5].RunComd := FALSE;
   BenchUut4.mode := FALSE;
   BenchUut4.start := TRUE;
   BenchUut4.stop := FALSE;
   TraceIn_mode[15] := BenchUut4.mode;
   TraceIn_start[15] := BenchUut4.start;
   TraceIn_stop[15] := BenchUut4.stop;
   BenchUut4(pumpGroup := Binding_4_pumpGroup);
   TraceOut_pumpGroup_1_priority[15] := Binding_4_pumpGroup[1].priority;
   TraceOut_pumpGroup_1_selection[15] := Binding_4_pumpGroup[1].selection;
   TraceOut_pumpGroup_1_RunComd[15] := Binding_4_pumpGroup[1].RunComd;
   TraceOut_pumpGroup_2_priority[15] := Binding_4_pumpGroup[2].priority;
   TraceOut_pumpGroup_2_selection[15] := Binding_4_pumpGroup[2].selection;
   TraceOut_pumpGroup_2_RunComd[15] := Binding_4_pumpGroup[2].RunComd;
   TraceOut_pumpGroup_3_priority[15] := Binding_4_pumpGroup[3].priority;
   TraceOut_pumpGroup_3_selection[15] := Binding_4_pumpGroup[3].selection;
   TraceOut_pumpGroup_3_RunComd[15] := Binding_4_pumpGroup[3].RunComd;
   TraceOut_pumpGroup_4_priority[15] := Binding_4_pumpGroup[4].priority;
   TraceOut_pumpGroup_4_selection[15] := Binding_4_pumpGroup[4].selection;
   TraceOut_pumpGroup_4_RunComd[15] := Binding_4_pumpGroup[4].RunComd;
   TraceOut_pumpGroup_5_priority[15] := Binding_4_pumpGroup[5].priority;
   TraceOut_pumpGroup_5_selection[15] := Binding_4_pumpGroup[5].selection;
   TraceOut_pumpGroup_5_RunComd[15] := Binding_4_pumpGroup[5].RunComd;
   BenchCalls := BenchCalls + 1;
 16:
   Binding_4_pumpGroup[1].priority := INT#10;
   Binding_4_pumpGroup[1].selection := FALSE;
   Binding_4_pumpGroup[1].RunComd := FALSE;
   Binding_4_pumpGroup[2].priority := INT#20;
   Binding_4_pumpGroup[2].selection := TRUE;
   Binding_4_pumpGroup[2].RunComd := FALSE;
   Binding_4_pumpGroup[3].priority := INT#30;
   Binding_4_pumpGroup[3].selection := FALSE;
   Binding_4_pumpGroup[3].RunComd := FALSE;
   Binding_4_pumpGroup[4].priority := INT#40;
   Binding_4_pumpGroup[4].selection := FALSE;
   Binding_4_pumpGroup[4].RunComd := FALSE;
   Binding_4_pumpGroup[5].priority := INT#50;
   Binding_4_pumpGroup[5].selection := TRUE;
   Binding_4_pumpGroup[5].RunComd := FALSE;
   BenchUut4.mode := FALSE;
   BenchUut4.start := TRUE;
   BenchUut4.stop := FALSE;
   TraceIn_mode[16] := BenchUut4.mode;
   TraceIn_start[16] := BenchUut4.start;
   TraceIn_stop[16] := BenchUut4.stop;
   BenchUut4(pumpGroup := Binding_4_pumpGroup);
   TraceOut_pumpGroup_1_priority[16] := Binding_4_pumpGroup[1].priority;
   TraceOut_pumpGroup_1_selection[16] := Binding_4_pumpGroup[1].selection;
   TraceOut_pumpGroup_1_RunComd[16] := Binding_4_pumpGroup[1].RunComd;
   TraceOut_pumpGroup_2_priority[16] := Binding_4_pumpGroup[2].priority;
   TraceOut_pumpGroup_2_selection[16] := Binding_4_pumpGroup[2].selection;
   TraceOut_pumpGroup_2_RunComd[16] := Binding_4_pumpGroup[2].RunComd;
   TraceOut_pumpGroup_3_priority[16] := Binding_4_pumpGroup[3].priority;
   TraceOut_pumpGroup_3_selection[16] := Binding_4_pumpGroup[3].selection;
   TraceOut_pumpGroup_3_RunComd[16] := Binding_4_pumpGroup[3].RunComd;
   TraceOut_pumpGroup_4_priority[16] := Binding_4_pumpGroup[4].priority;
   TraceOut_pumpGroup_4_selection[16] := Binding_4_pumpGroup[4].selection;
   TraceOut_pumpGroup_4_RunComd[16] := Binding_4_pumpGroup[4].RunComd;
   TraceOut_pumpGroup_5_priority[16] := Binding_4_pumpGroup[5].priority;
   TraceOut_pumpGroup_5_selection[16] := Binding_4_pumpGroup[5].selection;
   TraceOut_pumpGroup_5_RunComd[16] := Binding_4_pumpGroup[5].RunComd;
   BenchCalls := BenchCalls + 1;
 17:
   Binding_4_pumpGroup[1].priority := INT#10;
   Binding_4_pumpGroup[1].selection := FALSE;
   Binding_4_pumpGroup[1].RunComd := FALSE;
   Binding_4_pumpGroup[2].priority := INT#20;
   Binding_4_pumpGroup[2].selection := FALSE;
   Binding_4_pumpGroup[2].RunComd := TRUE;
   Binding_4_pumpGroup[3].priority := INT#30;
   Binding_4_pumpGroup[3].selection := FALSE;
   Binding_4_pumpGroup[3].RunComd := FALSE;
   Binding_4_pumpGroup[4].priority := INT#40;
   Binding_4_pumpGroup[4].selection := TRUE;
   Binding_4_pumpGroup[4].RunComd := FALSE;
   Binding_4_pumpGroup[5].priority := INT#50;
   Binding_4_pumpGroup[5].selection := FALSE;
   Binding_4_pumpGroup[5].RunComd := TRUE;
   BenchUut4.mode := FALSE;
   BenchUut4.start := FALSE;
   BenchUut4.stop := FALSE;
   TraceIn_mode[17] := BenchUut4.mode;
   TraceIn_start[17] := BenchUut4.start;
   TraceIn_stop[17] := BenchUut4.stop;
   BenchUut4(pumpGroup := Binding_4_pumpGroup);
   TraceOut_pumpGroup_1_priority[17] := Binding_4_pumpGroup[1].priority;
   TraceOut_pumpGroup_1_selection[17] := Binding_4_pumpGroup[1].selection;
   TraceOut_pumpGroup_1_RunComd[17] := Binding_4_pumpGroup[1].RunComd;
   TraceOut_pumpGroup_2_priority[17] := Binding_4_pumpGroup[2].priority;
   TraceOut_pumpGroup_2_selection[17] := Binding_4_pumpGroup[2].selection;
   TraceOut_pumpGroup_2_RunComd[17] := Binding_4_pumpGroup[2].RunComd;
   TraceOut_pumpGroup_3_priority[17] := Binding_4_pumpGroup[3].priority;
   TraceOut_pumpGroup_3_selection[17] := Binding_4_pumpGroup[3].selection;
   TraceOut_pumpGroup_3_RunComd[17] := Binding_4_pumpGroup[3].RunComd;
   TraceOut_pumpGroup_4_priority[17] := Binding_4_pumpGroup[4].priority;
   TraceOut_pumpGroup_4_selection[17] := Binding_4_pumpGroup[4].selection;
   TraceOut_pumpGroup_4_RunComd[17] := Binding_4_pumpGroup[4].RunComd;
   TraceOut_pumpGroup_5_priority[17] := Binding_4_pumpGroup[5].priority;
   TraceOut_pumpGroup_5_selection[17] := Binding_4_pumpGroup[5].selection;
   TraceOut_pumpGroup_5_RunComd[17] := Binding_4_pumpGroup[5].RunComd;
   BenchCalls := BenchCalls + 1;
 18:
   Binding_4_pumpGroup[1].priority := INT#10;
   Binding_4_pumpGroup[1].selection := FALSE;
   Binding_4_pumpGroup[1].RunComd := FALSE;
   Binding_4_pumpGroup[2].priority := INT#20;
   Binding_4_pumpGroup[2].selection := FALSE;
   Binding_4_pumpGroup[2].RunComd := TRUE;
   Binding_4_pumpGroup[3].priority := INT#30;
   Binding_4_pumpGroup[3].selection := FALSE;
   Binding_4_pumpGroup[3].RunComd := FALSE;
   Binding_4_pumpGroup[4].priority := INT#40;
   Binding_4_pumpGroup[4].selection := TRUE;
   Binding_4_pumpGroup[4].RunComd := FALSE;
   Binding_4_pumpGroup[5].priority := INT#50;
   Binding_4_pumpGroup[5].selection := FALSE;
   Binding_4_pumpGroup[5].RunComd := TRUE;
   BenchUut4.mode := FALSE;
   BenchUut4.start := TRUE;
   BenchUut4.stop := FALSE;
   TraceIn_mode[18] := BenchUut4.mode;
   TraceIn_start[18] := BenchUut4.start;
   TraceIn_stop[18] := BenchUut4.stop;
   BenchUut4(pumpGroup := Binding_4_pumpGroup);
   TraceOut_pumpGroup_1_priority[18] := Binding_4_pumpGroup[1].priority;
   TraceOut_pumpGroup_1_selection[18] := Binding_4_pumpGroup[1].selection;
   TraceOut_pumpGroup_1_RunComd[18] := Binding_4_pumpGroup[1].RunComd;
   TraceOut_pumpGroup_2_priority[18] := Binding_4_pumpGroup[2].priority;
   TraceOut_pumpGroup_2_selection[18] := Binding_4_pumpGroup[2].selection;
   TraceOut_pumpGroup_2_RunComd[18] := Binding_4_pumpGroup[2].RunComd;
   TraceOut_pumpGroup_3_priority[18] := Binding_4_pumpGroup[3].priority;
   TraceOut_pumpGroup_3_selection[18] := Binding_4_pumpGroup[3].selection;
   TraceOut_pumpGroup_3_RunComd[18] := Binding_4_pumpGroup[3].RunComd;
   TraceOut_pumpGroup_4_priority[18] := Binding_4_pumpGroup[4].priority;
   TraceOut_pumpGroup_4_selection[18] := Binding_4_pumpGroup[4].selection;
   TraceOut_pumpGroup_4_RunComd[18] := Binding_4_pumpGroup[4].RunComd;
   TraceOut_pumpGroup_5_priority[18] := Binding_4_pumpGroup[5].priority;
   TraceOut_pumpGroup_5_selection[18] := Binding_4_pumpGroup[5].selection;
   TraceOut_pumpGroup_5_RunComd[18] := Binding_4_pumpGroup[5].RunComd;
   BenchCalls := BenchCalls + 1;
 19:
   Binding_4_pumpGroup[1].priority := INT#10;
   Binding_4_pumpGroup[1].selection := FALSE;
   Binding_4_pumpGroup[1].RunComd := FALSE;
   Binding_4_pumpGroup[2].priority := INT#20;
   Binding_4_pumpGroup[2].selection := FALSE;
   Binding_4_pumpGroup[2].RunComd := TRUE;
   Binding_4_pumpGroup[3].priority := INT#30;
   Binding_4_pumpGroup[3].selection := FALSE;
   Binding_4_pumpGroup[3].RunComd := FALSE;
   Binding_4_pumpGroup[4].priority := INT#40;
   Binding_4_pumpGroup[4].selection := TRUE;
   Binding_4_pumpGroup[4].RunComd := FALSE;
   Binding_4_pumpGroup[5].priority := INT#50;
   Binding_4_pumpGroup[5].selection := FALSE;
   Binding_4_pumpGroup[5].RunComd := TRUE;
   BenchUut4.mode := TRUE;
   BenchUut4.start := TRUE;
   BenchUut4.stop := FALSE;
   TraceIn_mode[19] := BenchUut4.mode;
   TraceIn_start[19] := BenchUut4.start;
   TraceIn_stop[19] := BenchUut4.stop;
   BenchUut4(pumpGroup := Binding_4_pumpGroup);
   TraceOut_pumpGroup_1_priority[19] := Binding_4_pumpGroup[1].priority;
   TraceOut_pumpGroup_1_selection[19] := Binding_4_pumpGroup[1].selection;
   TraceOut_pumpGroup_1_RunComd[19] := Binding_4_pumpGroup[1].RunComd;
   TraceOut_pumpGroup_2_priority[19] := Binding_4_pumpGroup[2].priority;
   TraceOut_pumpGroup_2_selection[19] := Binding_4_pumpGroup[2].selection;
   TraceOut_pumpGroup_2_RunComd[19] := Binding_4_pumpGroup[2].RunComd;
   TraceOut_pumpGroup_3_priority[19] := Binding_4_pumpGroup[3].priority;
   TraceOut_pumpGroup_3_selection[19] := Binding_4_pumpGroup[3].selection;
   TraceOut_pumpGroup_3_RunComd[19] := Binding_4_pumpGroup[3].RunComd;
   TraceOut_pumpGroup_4_priority[19] := Binding_4_pumpGroup[4].priority;
   TraceOut_pumpGroup_4_selection[19] := Binding_4_pumpGroup[4].selection;
   TraceOut_pumpGroup_4_RunComd[19] := Binding_4_pumpGroup[4].RunComd;
   TraceOut_pumpGroup_5_priority[19] := Binding_4_pumpGroup[5].priority;
   TraceOut_pumpGroup_5_selection[19] := Binding_4_pumpGroup[5].selection;
   TraceOut_pumpGroup_5_RunComd[19] := Binding_4_pumpGroup[5].RunComd;
   BenchCalls := BenchCalls + 1;
 20:
   Binding_4_pumpGroup[1].priority := INT#10;
   Binding_4_pumpGroup[1].selection := FALSE;
   Binding_4_pumpGroup[1].RunComd := FALSE;
   Binding_4_pumpGroup[2].priority := INT#20;
   Binding_4_pumpGroup[2].selection := FALSE;
   Binding_4_pumpGroup[2].RunComd := TRUE;
   Binding_4_pumpGroup[3].priority := INT#30;
   Binding_4_pumpGroup[3].selection := FALSE;
   Binding_4_pumpGroup[3].RunComd := FALSE;
   Binding_4_pumpGroup[4].priority := INT#40;
   Binding_4_pumpGroup[4].selection := TRUE;
   Binding_4_pumpGroup[4].RunComd := FALSE;
   Binding_4_pumpGroup[5].priority := INT#50;
   Binding_4_pumpGroup[5].selection := FALSE;
   Binding_4_pumpGroup[5].RunComd := TRUE;
   BenchUut4.mode := FALSE;
   BenchUut4.start := TRUE;
   BenchUut4.stop := FALSE;
   TraceIn_mode[20] := BenchUut4.mode;
   TraceIn_start[20] := BenchUut4.start;
   TraceIn_stop[20] := BenchUut4.stop;
   BenchUut4(pumpGroup := Binding_4_pumpGroup);
   TraceOut_pumpGroup_1_priority[20] := Binding_4_pumpGroup[1].priority;
   TraceOut_pumpGroup_1_selection[20] := Binding_4_pumpGroup[1].selection;
   TraceOut_pumpGroup_1_RunComd[20] := Binding_4_pumpGroup[1].RunComd;
   TraceOut_pumpGroup_2_priority[20] := Binding_4_pumpGroup[2].priority;
   TraceOut_pumpGroup_2_selection[20] := Binding_4_pumpGroup[2].selection;
   TraceOut_pumpGroup_2_RunComd[20] := Binding_4_pumpGroup[2].RunComd;
   TraceOut_pumpGroup_3_priority[20] := Binding_4_pumpGroup[3].priority;
   TraceOut_pumpGroup_3_selection[20] := Binding_4_pumpGroup[3].selection;
   TraceOut_pumpGroup_3_RunComd[20] := Binding_4_pumpGroup[3].RunComd;
   TraceOut_pumpGroup_4_priority[20] := Binding_4_pumpGroup[4].priority;
   TraceOut_pumpGroup_4_selection[20] := Binding_4_pumpGroup[4].selection;
   TraceOut_pumpGroup_4_RunComd[20] := Binding_4_pumpGroup[4].RunComd;
   TraceOut_pumpGroup_5_priority[20] := Binding_4_pumpGroup[5].priority;
   TraceOut_pumpGroup_5_selection[20] := Binding_4_pumpGroup[5].selection;
   TraceOut_pumpGroup_5_RunComd[20] := Binding_4_pumpGroup[5].RunComd;
   BenchCalls := BenchCalls + 1;
 21:
   Binding_4_pumpGroup[1].priority := INT#10;
   Binding_4_pumpGroup[1].selection := FALSE;
   Binding_4_pumpGroup[1].RunComd := FALSE;
   Binding_4_pumpGroup[2].priority := INT#20;
   Binding_4_pumpGroup[2].selection := FALSE;
   Binding_4_pumpGroup[2].RunComd := TRUE;
   Binding_4_pumpGroup[3].priority := INT#30;
   Binding_4_pumpGroup[3].selection := FALSE;
   Binding_4_pumpGroup[3].RunComd := FALSE;
   Binding_4_pumpGroup[4].priority := INT#40;
   Binding_4_pumpGroup[4].selection := TRUE;
   Binding_4_pumpGroup[4].RunComd := FALSE;
   Binding_4_pumpGroup[5].priority := INT#50;
   Binding_4_pumpGroup[5].selection := FALSE;
   Binding_4_pumpGroup[5].RunComd := TRUE;
   BenchUut4.mode := FALSE;
   BenchUut4.start := TRUE;
   BenchUut4.stop := TRUE;
   TraceIn_mode[21] := BenchUut4.mode;
   TraceIn_start[21] := BenchUut4.start;
   TraceIn_stop[21] := BenchUut4.stop;
   BenchUut4(pumpGroup := Binding_4_pumpGroup);
   TraceOut_pumpGroup_1_priority[21] := Binding_4_pumpGroup[1].priority;
   TraceOut_pumpGroup_1_selection[21] := Binding_4_pumpGroup[1].selection;
   TraceOut_pumpGroup_1_RunComd[21] := Binding_4_pumpGroup[1].RunComd;
   TraceOut_pumpGroup_2_priority[21] := Binding_4_pumpGroup[2].priority;
   TraceOut_pumpGroup_2_selection[21] := Binding_4_pumpGroup[2].selection;
   TraceOut_pumpGroup_2_RunComd[21] := Binding_4_pumpGroup[2].RunComd;
   TraceOut_pumpGroup_3_priority[21] := Binding_4_pumpGroup[3].priority;
   TraceOut_pumpGroup_3_selection[21] := Binding_4_pumpGroup[3].selection;
   TraceOut_pumpGroup_3_RunComd[21] := Binding_4_pumpGroup[3].RunComd;
   TraceOut_pumpGroup_4_priority[21] := Binding_4_pumpGroup[4].priority;
   TraceOut_pumpGroup_4_selection[21] := Binding_4_pumpGroup[4].selection;
   TraceOut_pumpGroup_4_RunComd[21] := Binding_4_pumpGroup[4].RunComd;
   TraceOut_pumpGroup_5_priority[21] := Binding_4_pumpGroup[5].priority;
   TraceOut_pumpGroup_5_selection[21] := Binding_4_pumpGroup[5].selection;
   TraceOut_pumpGroup_5_RunComd[21] := Binding_4_pumpGroup[5].RunComd;
   BenchCalls := BenchCalls + 1;
 22:
   Binding_5_pumpGroup[1].priority := INT#-5;
   Binding_5_pumpGroup[1].selection := FALSE;
   Binding_5_pumpGroup[1].RunComd := FALSE;
   Binding_5_pumpGroup[2].priority := INT#-1;
   Binding_5_pumpGroup[2].selection := FALSE;
   Binding_5_pumpGroup[2].RunComd := FALSE;
   Binding_5_pumpGroup[3].priority := INT#0;
   Binding_5_pumpGroup[3].selection := FALSE;
   Binding_5_pumpGroup[3].RunComd := FALSE;
   Binding_5_pumpGroup[4].priority := INT#-5;
   Binding_5_pumpGroup[4].selection := TRUE;
   Binding_5_pumpGroup[4].RunComd := FALSE;
   Binding_5_pumpGroup[5].priority := INT#-10;
   Binding_5_pumpGroup[5].selection := TRUE;
   Binding_5_pumpGroup[5].RunComd := FALSE;
   BenchUut5.mode := TRUE;
   BenchUut5.start := TRUE;
   BenchUut5.stop := FALSE;
   TraceIn_mode[22] := BenchUut5.mode;
   TraceIn_start[22] := BenchUut5.start;
   TraceIn_stop[22] := BenchUut5.stop;
   BenchUut5(pumpGroup := Binding_5_pumpGroup);
   TraceOut_pumpGroup_1_priority[22] := Binding_5_pumpGroup[1].priority;
   TraceOut_pumpGroup_1_selection[22] := Binding_5_pumpGroup[1].selection;
   TraceOut_pumpGroup_1_RunComd[22] := Binding_5_pumpGroup[1].RunComd;
   TraceOut_pumpGroup_2_priority[22] := Binding_5_pumpGroup[2].priority;
   TraceOut_pumpGroup_2_selection[22] := Binding_5_pumpGroup[2].selection;
   TraceOut_pumpGroup_2_RunComd[22] := Binding_5_pumpGroup[2].RunComd;
   TraceOut_pumpGroup_3_priority[22] := Binding_5_pumpGroup[3].priority;
   TraceOut_pumpGroup_3_selection[22] := Binding_5_pumpGroup[3].selection;
   TraceOut_pumpGroup_3_RunComd[22] := Binding_5_pumpGroup[3].RunComd;
   TraceOut_pumpGroup_4_priority[22] := Binding_5_pumpGroup[4].priority;
   TraceOut_pumpGroup_4_selection[22] := Binding_5_pumpGroup[4].selection;
   TraceOut_pumpGroup_4_RunComd[22] := Binding_5_pumpGroup[4].RunComd;
   TraceOut_pumpGroup_5_priority[22] := Binding_5_pumpGroup[5].priority;
   TraceOut_pumpGroup_5_selection[22] := Binding_5_pumpGroup[5].selection;
   TraceOut_pumpGroup_5_RunComd[22] := Binding_5_pumpGroup[5].RunComd;
   BenchCalls := BenchCalls + 1;
 23:
   Binding_5_pumpGroup[1].priority := INT#-3;
   Binding_5_pumpGroup[1].selection := FALSE;
   Binding_5_pumpGroup[1].RunComd := TRUE;
   Binding_5_pumpGroup[2].priority := INT#-3;
   Binding_5_pumpGroup[2].selection := FALSE;
   Binding_5_pumpGroup[2].RunComd := TRUE;
   Binding_5_pumpGroup[3].priority := INT#-3;
   Binding_5_pumpGroup[3].selection := FALSE;
   Binding_5_pumpGroup[3].RunComd := TRUE;
   Binding_5_pumpGroup[4].priority := INT#-3;
   Binding_5_pumpGroup[4].selection := TRUE;
   Binding_5_pumpGroup[4].RunComd := FALSE;
   Binding_5_pumpGroup[5].priority := INT#-3;
   Binding_5_pumpGroup[5].selection := TRUE;
   Binding_5_pumpGroup[5].RunComd := FALSE;
   BenchUut5.mode := TRUE;
   BenchUut5.start := TRUE;
   BenchUut5.stop := FALSE;
   TraceIn_mode[23] := BenchUut5.mode;
   TraceIn_start[23] := BenchUut5.start;
   TraceIn_stop[23] := BenchUut5.stop;
   BenchUut5(pumpGroup := Binding_5_pumpGroup);
   TraceOut_pumpGroup_1_priority[23] := Binding_5_pumpGroup[1].priority;
   TraceOut_pumpGroup_1_selection[23] := Binding_5_pumpGroup[1].selection;
   TraceOut_pumpGroup_1_RunComd[23] := Binding_5_pumpGroup[1].RunComd;
   TraceOut_pumpGroup_2_priority[23] := Binding_5_pumpGroup[2].priority;
   TraceOut_pumpGroup_2_selection[23] := Binding_5_pumpGroup[2].selection;
   TraceOut_pumpGroup_2_RunComd[23] := Binding_5_pumpGroup[2].RunComd;
   TraceOut_pumpGroup_3_priority[23] := Binding_5_pumpGroup[3].priority;
   TraceOut_pumpGroup_3_selection[23] := Binding_5_pumpGroup[3].selection;
   TraceOut_pumpGroup_3_RunComd[23] := Binding_5_pumpGroup[3].RunComd;
   TraceOut_pumpGroup_4_priority[23] := Binding_5_pumpGroup[4].priority;
   TraceOut_pumpGroup_4_selection[23] := Binding_5_pumpGroup[4].selection;
   TraceOut_pumpGroup_4_RunComd[23] := Binding_5_pumpGroup[4].RunComd;
   TraceOut_pumpGroup_5_priority[23] := Binding_5_pumpGroup[5].priority;
   TraceOut_pumpGroup_5_selection[23] := Binding_5_pumpGroup[5].selection;
   TraceOut_pumpGroup_5_RunComd[23] := Binding_5_pumpGroup[5].RunComd;
   BenchCalls := BenchCalls + 1;
 24:
   Binding_5_pumpGroup[1].priority := INT#100;
   Binding_5_pumpGroup[1].selection := FALSE;
   Binding_5_pumpGroup[1].RunComd := TRUE;
   Binding_5_pumpGroup[2].priority := INT#90;
   Binding_5_pumpGroup[2].selection := FALSE;
   Binding_5_pumpGroup[2].RunComd := TRUE;
   Binding_5_pumpGroup[3].priority := INT#80;
   Binding_5_pumpGroup[3].selection := FALSE;
   Binding_5_pumpGroup[3].RunComd := TRUE;
   Binding_5_pumpGroup[4].priority := INT#70;
   Binding_5_pumpGroup[4].selection := FALSE;
   Binding_5_pumpGroup[4].RunComd := FALSE;
   Binding_5_pumpGroup[5].priority := INT#60;
   Binding_5_pumpGroup[5].selection := FALSE;
   Binding_5_pumpGroup[5].RunComd := FALSE;
   BenchUut5.mode := FALSE;
   BenchUut5.start := TRUE;
   BenchUut5.stop := FALSE;
   TraceIn_mode[24] := BenchUut5.mode;
   TraceIn_start[24] := BenchUut5.start;
   TraceIn_stop[24] := BenchUut5.stop;
   BenchUut5(pumpGroup := Binding_5_pumpGroup);
   TraceOut_pumpGroup_1_priority[24] := Binding_5_pumpGroup[1].priority;
   TraceOut_pumpGroup_1_selection[24] := Binding_5_pumpGroup[1].selection;
   TraceOut_pumpGroup_1_RunComd[24] := Binding_5_pumpGroup[1].RunComd;
   TraceOut_pumpGroup_2_priority[24] := Binding_5_pumpGroup[2].priority;
   TraceOut_pumpGroup_2_selection[24] := Binding_5_pumpGroup[2].selection;
   TraceOut_pumpGroup_2_RunComd[24] := Binding_5_pumpGroup[2].RunComd;
   TraceOut_pumpGroup_3_priority[24] := Binding_5_pumpGroup[3].priority;
   TraceOut_pumpGroup_3_selection[24] := Binding_5_pumpGroup[3].selection;
   TraceOut_pumpGroup_3_RunComd[24] := Binding_5_pumpGroup[3].RunComd;
   TraceOut_pumpGroup_4_priority[24] := Binding_5_pumpGroup[4].priority;
   TraceOut_pumpGroup_4_selection[24] := Binding_5_pumpGroup[4].selection;
   TraceOut_pumpGroup_4_RunComd[24] := Binding_5_pumpGroup[4].RunComd;
   TraceOut_pumpGroup_5_priority[24] := Binding_5_pumpGroup[5].priority;
   TraceOut_pumpGroup_5_selection[24] := Binding_5_pumpGroup[5].selection;
   TraceOut_pumpGroup_5_RunComd[24] := Binding_5_pumpGroup[5].RunComd;
   BenchCalls := BenchCalls + 1;
 25:
   Binding_5_pumpGroup[1].priority := INT#100;
   Binding_5_pumpGroup[1].selection := FALSE;
   Binding_5_pumpGroup[1].RunComd := FALSE;
   Binding_5_pumpGroup[2].priority := INT#90;
   Binding_5_pumpGroup[2].selection := FALSE;
   Binding_5_pumpGroup[2].RunComd := FALSE;
   Binding_5_pumpGroup[3].priority := INT#80;
   Binding_5_pumpGroup[3].selection := TRUE;
   Binding_5_pumpGroup[3].RunComd := FALSE;
   Binding_5_pumpGroup[4].priority := INT#70;
   Binding_5_pumpGroup[4].selection := FALSE;
   Binding_5_pumpGroup[4].RunComd := FALSE;
   Binding_5_pumpGroup[5].priority := INT#60;
   Binding_5_pumpGroup[5].selection := TRUE;
   Binding_5_pumpGroup[5].RunComd := FALSE;
   BenchUut5.mode := FALSE;
   BenchUut5.start := TRUE;
   BenchUut5.stop := FALSE;
   TraceIn_mode[25] := BenchUut5.mode;
   TraceIn_start[25] := BenchUut5.start;
   TraceIn_stop[25] := BenchUut5.stop;
   BenchUut5(pumpGroup := Binding_5_pumpGroup);
   TraceOut_pumpGroup_1_priority[25] := Binding_5_pumpGroup[1].priority;
   TraceOut_pumpGroup_1_selection[25] := Binding_5_pumpGroup[1].selection;
   TraceOut_pumpGroup_1_RunComd[25] := Binding_5_pumpGroup[1].RunComd;
   TraceOut_pumpGroup_2_priority[25] := Binding_5_pumpGroup[2].priority;
   TraceOut_pumpGroup_2_selection[25] := Binding_5_pumpGroup[2].selection;
   TraceOut_pumpGroup_2_RunComd[25] := Binding_5_pumpGroup[2].RunComd;
   TraceOut_pumpGroup_3_priority[25] := Binding_5_pumpGroup[3].priority;
   TraceOut_pumpGroup_3_selection[25] := Binding_5_pumpGroup[3].selection;
   TraceOut_pumpGroup_3_RunComd[25] := Binding_5_pumpGroup[3].RunComd;
   TraceOut_pumpGroup_4_priority[25] := Binding_5_pumpGroup[4].priority;
   TraceOut_pumpGroup_4_selection[25] := Binding_5_pumpGroup[4].selection;
   TraceOut_pumpGroup_4_RunComd[25] := Binding_5_pumpGroup[4].RunComd;
   TraceOut_pumpGroup_5_priority[25] := Binding_5_pumpGroup[5].priority;
   TraceOut_pumpGroup_5_selection[25] := Binding_5_pumpGroup[5].selection;
   TraceOut_pumpGroup_5_RunComd[25] := Binding_5_pumpGroup[5].RunComd;
   BenchCalls := BenchCalls + 1;
 26:
   Binding_6_pumpGroup[1].priority := INT#50;
   Binding_6_pumpGroup[1].selection := TRUE;
   Binding_6_pumpGroup[1].RunComd := FALSE;
   Binding_6_pumpGroup[2].priority := INT#10;
   Binding_6_pumpGroup[2].selection := TRUE;
   Binding_6_pumpGroup[2].RunComd := FALSE;
   Binding_6_pumpGroup[3].priority := INT#40;
   Binding_6_pumpGroup[3].selection := TRUE;
   Binding_6_pumpGroup[3].RunComd := FALSE;
   Binding_6_pumpGroup[4].priority := INT#20;
   Binding_6_pumpGroup[4].selection := TRUE;
   Binding_6_pumpGroup[4].RunComd := FALSE;
   Binding_6_pumpGroup[5].priority := INT#25;
   Binding_6_pumpGroup[5].selection := TRUE;
   Binding_6_pumpGroup[5].RunComd := FALSE;
   BenchUut6.mode := TRUE;
   BenchUut6.start := TRUE;
   BenchUut6.stop := FALSE;
   TraceIn_mode[26] := BenchUut6.mode;
   TraceIn_start[26] := BenchUut6.start;
   TraceIn_stop[26] := BenchUut6.stop;
   BenchUut6(pumpGroup := Binding_6_pumpGroup);
   TraceOut_pumpGroup_1_priority[26] := Binding_6_pumpGroup[1].priority;
   TraceOut_pumpGroup_1_selection[26] := Binding_6_pumpGroup[1].selection;
   TraceOut_pumpGroup_1_RunComd[26] := Binding_6_pumpGroup[1].RunComd;
   TraceOut_pumpGroup_2_priority[26] := Binding_6_pumpGroup[2].priority;
   TraceOut_pumpGroup_2_selection[26] := Binding_6_pumpGroup[2].selection;
   TraceOut_pumpGroup_2_RunComd[26] := Binding_6_pumpGroup[2].RunComd;
   TraceOut_pumpGroup_3_priority[26] := Binding_6_pumpGroup[3].priority;
   TraceOut_pumpGroup_3_selection[26] := Binding_6_pumpGroup[3].selection;
   TraceOut_pumpGroup_3_RunComd[26] := Binding_6_pumpGroup[3].RunComd;
   TraceOut_pumpGroup_4_priority[26] := Binding_6_pumpGroup[4].priority;
   TraceOut_pumpGroup_4_selection[26] := Binding_6_pumpGroup[4].selection;
   TraceOut_pumpGroup_4_RunComd[26] := Binding_6_pumpGroup[4].RunComd;
   TraceOut_pumpGroup_5_priority[26] := Binding_6_pumpGroup[5].priority;
   TraceOut_pumpGroup_5_selection[26] := Binding_6_pumpGroup[5].selection;
   TraceOut_pumpGroup_5_RunComd[26] := Binding_6_pumpGroup[5].RunComd;
   BenchCalls := BenchCalls + 1;
 27:
   Binding_6_pumpGroup[1].priority := INT#1;
   Binding_6_pumpGroup[1].selection := TRUE;
   Binding_6_pumpGroup[1].RunComd := TRUE;
   Binding_6_pumpGroup[2].priority := INT#99;
   Binding_6_pumpGroup[2].selection := TRUE;
   Binding_6_pumpGroup[2].RunComd := FALSE;
   Binding_6_pumpGroup[3].priority := INT#2;
   Binding_6_pumpGroup[3].selection := FALSE;
   Binding_6_pumpGroup[3].RunComd := TRUE;
   Binding_6_pumpGroup[4].priority := INT#88;
   Binding_6_pumpGroup[4].selection := FALSE;
   Binding_6_pumpGroup[4].RunComd := FALSE;
   Binding_6_pumpGroup[5].priority := INT#77;
   Binding_6_pumpGroup[5].selection := FALSE;
   Binding_6_pumpGroup[5].RunComd := TRUE;
   BenchUut6.mode := FALSE;
   BenchUut6.start := FALSE;
   BenchUut6.stop := FALSE;
   TraceIn_mode[27] := BenchUut6.mode;
   TraceIn_start[27] := BenchUut6.start;
   TraceIn_stop[27] := BenchUut6.stop;
   BenchUut6(pumpGroup := Binding_6_pumpGroup);
   TraceOut_pumpGroup_1_priority[27] := Binding_6_pumpGroup[1].priority;
   TraceOut_pumpGroup_1_selection[27] := Binding_6_pumpGroup[1].selection;
   TraceOut_pumpGroup_1_RunComd[27] := Binding_6_pumpGroup[1].RunComd;
   TraceOut_pumpGroup_2_priority[27] := Binding_6_pumpGroup[2].priority;
   TraceOut_pumpGroup_2_selection[27] := Binding_6_pumpGroup[2].selection;
   TraceOut_pumpGroup_2_RunComd[27] := Binding_6_pumpGroup[2].RunComd;
   TraceOut_pumpGroup_3_priority[27] := Binding_6_pumpGroup[3].priority;
   TraceOut_pumpGroup_3_selection[27] := Binding_6_pumpGroup[3].selection;
   TraceOut_pumpGroup_3_RunComd[27] := Binding_6_pumpGroup[3].RunComd;
   TraceOut_pumpGroup_4_priority[27] := Binding_6_pumpGroup[4].priority;
   TraceOut_pumpGroup_4_selection[27] := Binding_6_pumpGroup[4].selection;
   TraceOut_pumpGroup_4_RunComd[27] := Binding_6_pumpGroup[4].RunComd;
   TraceOut_pumpGroup_5_priority[27] := Binding_6_pumpGroup[5].priority;
   TraceOut_pumpGroup_5_selection[27] := Binding_6_pumpGroup[5].selection;
   TraceOut_pumpGroup_5_RunComd[27] := Binding_6_pumpGroup[5].RunComd;
   BenchCalls := BenchCalls + 1;
 28:
   Binding_6_pumpGroup[1].priority := INT#1;
   Binding_6_pumpGroup[1].selection := TRUE;
   Binding_6_pumpGroup[1].RunComd := TRUE;
   Binding_6_pumpGroup[2].priority := INT#99;
   Binding_6_pumpGroup[2].selection := TRUE;
   Binding_6_pumpGroup[2].RunComd := FALSE;
   Binding_6_pumpGroup[3].priority := INT#2;
   Binding_6_pumpGroup[3].selection := FALSE;
   Binding_6_pumpGroup[3].RunComd := TRUE;
   Binding_6_pumpGroup[4].priority := INT#88;
   Binding_6_pumpGroup[4].selection := FALSE;
   Binding_6_pumpGroup[4].RunComd := FALSE;
   Binding_6_pumpGroup[5].priority := INT#77;
   Binding_6_pumpGroup[5].selection := FALSE;
   Binding_6_pumpGroup[5].RunComd := TRUE;
   BenchUut6.mode := FALSE;
   BenchUut6.start := TRUE;
   BenchUut6.stop := FALSE;
   TraceIn_mode[28] := BenchUut6.mode;
   TraceIn_start[28] := BenchUut6.start;
   TraceIn_stop[28] := BenchUut6.stop;
   BenchUut6(pumpGroup := Binding_6_pumpGroup);
   TraceOut_pumpGroup_1_priority[28] := Binding_6_pumpGroup[1].priority;
   TraceOut_pumpGroup_1_selection[28] := Binding_6_pumpGroup[1].selection;
   TraceOut_pumpGroup_1_RunComd[28] := Binding_6_pumpGroup[1].RunComd;
   TraceOut_pumpGroup_2_priority[28] := Binding_6_pumpGroup[2].priority;
   TraceOut_pumpGroup_2_selection[28] := Binding_6_pumpGroup[2].selection;
   TraceOut_pumpGroup_2_RunComd[28] := Binding_6_pumpGroup[2].RunComd;
   TraceOut_pumpGroup_3_priority[28] := Binding_6_pumpGroup[3].priority;
   TraceOut_pumpGroup_3_selection[28] := Binding_6_pumpGroup[3].selection;
   TraceOut_pumpGroup_3_RunComd[28] := Binding_6_pumpGroup[3].RunComd;
   TraceOut_pumpGroup_4_priority[28] := Binding_6_pumpGroup[4].priority;
   TraceOut_pumpGroup_4_selection[28] := Binding_6_pumpGroup[4].selection;
   TraceOut_pumpGroup_4_RunComd[28] := Binding_6_pumpGroup[4].RunComd;
   TraceOut_pumpGroup_5_priority[28] := Binding_6_pumpGroup[5].priority;
   TraceOut_pumpGroup_5_selection[28] := Binding_6_pumpGroup[5].selection;
   TraceOut_pumpGroup_5_RunComd[28] := Binding_6_pumpGroup[5].RunComd;
   BenchCalls := BenchCalls + 1;
 29:
   Binding_6_pumpGroup[1].priority := INT#1;
   Binding_6_pumpGroup[1].selection := TRUE;
   Binding_6_pumpGroup[1].RunComd := TRUE;
   Binding_6_pumpGroup[2].priority := INT#2;
   Binding_6_pumpGroup[2].selection := TRUE;
   Binding_6_pumpGroup[2].RunComd := TRUE;
   Binding_6_pumpGroup[3].priority := INT#3;
   Binding_6_pumpGroup[3].selection := TRUE;
   Binding_6_pumpGroup[3].RunComd := FALSE;
   Binding_6_pumpGroup[4].priority := INT#4;
   Binding_6_pumpGroup[4].selection := FALSE;
   Binding_6_pumpGroup[4].RunComd := FALSE;
   Binding_6_pumpGroup[5].priority := INT#5;
   Binding_6_pumpGroup[5].selection := FALSE;
   Binding_6_pumpGroup[5].RunComd := FALSE;
   BenchUut6.mode := TRUE;
   BenchUut6.start := TRUE;
   BenchUut6.stop := TRUE;
   TraceIn_mode[29] := BenchUut6.mode;
   TraceIn_start[29] := BenchUut6.start;
   TraceIn_stop[29] := BenchUut6.stop;
   BenchUut6(pumpGroup := Binding_6_pumpGroup);
   TraceOut_pumpGroup_1_priority[29] := Binding_6_pumpGroup[1].priority;
   TraceOut_pumpGroup_1_selection[29] := Binding_6_pumpGroup[1].selection;
   TraceOut_pumpGroup_1_RunComd[29] := Binding_6_pumpGroup[1].RunComd;
   TraceOut_pumpGroup_2_priority[29] := Binding_6_pumpGroup[2].priority;
   TraceOut_pumpGroup_2_selection[29] := Binding_6_pumpGroup[2].selection;
   TraceOut_pumpGroup_2_RunComd[29] := Binding_6_pumpGroup[2].RunComd;
   TraceOut_pumpGroup_3_priority[29] := Binding_6_pumpGroup[3].priority;
   TraceOut_pumpGroup_3_selection[29] := Binding_6_pumpGroup[3].selection;
   TraceOut_pumpGroup_3_RunComd[29] := Binding_6_pumpGroup[3].RunComd;
   TraceOut_pumpGroup_4_priority[29] := Binding_6_pumpGroup[4].priority;
   TraceOut_pumpGroup_4_selection[29] := Binding_6_pumpGroup[4].selection;
   TraceOut_pumpGroup_4_RunComd[29] := Binding_6_pumpGroup[4].RunComd;
   TraceOut_pumpGroup_5_priority[29] := Binding_6_pumpGroup[5].priority;
   TraceOut_pumpGroup_5_selection[29] := Binding_6_pumpGroup[5].selection;
   TraceOut_pumpGroup_5_RunComd[29] := Binding_6_pumpGroup[5].RunComd;
   BenchCalls := BenchCalls + 1;
 END_CASE;
 BenchStep := BenchStep + 1;
 IF BenchStep >= 30 THEN BenchDone := TRUE; END_IF;
END_IF;
END_PROGRAM
